(* IEC 61131-3 sources: 2026_Projet_YGO_ExcavatriceDragage/ARCHIVES/Code/SUPERVISION, 3 files *)

(* ---- ST_Safety_Emergency_HmiCmd.st ---- *)
(* ==============================================================
   [IHM] ST_Safety_Emergency_HmiCmd -- Commandes IHM pour la chaine AU
   --------------------------------------------------------------
   Role : structure d'echange pour les commandes operateur
          de la chaine d'arret d'urgence (miroir ST_ModesCmd).
   Pattern : identique a GVL_IHM.Modes.Cmd dans le projet reel.
          L'IHM ecrit ces champs, le programme les consomme.
   ==============================================================
    Docs : DOC/AF/AF_Partie-01_Analyse_Fonctionnelle_v2.0.md
           DOC/AF/AF_Partie-07_Interface_IHM_v2.0.md
*)

TYPE ST_Safety_Emergency_HmiCmd :
STRUCT
    BtnEmergencyArming   : BOOL;   // Front demande rearmement contacteur
    BtnEmergencyCutOff   : BOOL;   // Niveau coupure IHM maintenue
    BtnFaultReset        : BOOL;   // Front acquittement defauts
END_STRUCT
END_TYPE

(* ---- ST_Safety_Emergency_HmiState.st ---- *)
(* ==============================================================
   [IHM] ST_Safety_Emergency_HmiState -- Retours d'etat IHM pour chaine AU
   --------------------------------------------------------------
   Role : structure d'echange pour les retours d'etat de la
          chaine d'arret d'urgence (miroir ST_ModesState).
   Pattern : identique a GVL_IHM.Modes.State dans le projet reel.
          Le programme ecrit ces champs, l'IHM les lit.
   ==============================================================
    Docs : DOC/AF/AF_Partie-01_Analyse_Fonctionnelle_v2.0.md
           DOC/AF/AF_Partie-07_Interface_IHM_v2.0.md
*)

TYPE ST_Safety_Emergency_HmiState :
STRUCT
    // [OK] Etats generaux
    ChainOk              : BOOL;   // Boucle AU fermee (saine)
    ContactorOk          : BOOL;   // Contacteur puissance engage
    PowerCutOffActive    : BOOL;   // Coupure puissance demandee par une safety metier

    // [AU] Sequence de rearmement
    Armable              : BOOL;   // Pret au rearmement (chain OK + pas de lockout + pas de defaut)
    ArmingBusy           : BOOL;   // Sequence armement en cours
    Step                 : INT;    // Etape sequence (0=IDLE, 1=TestA, 2=RestoreA, 3=TestB, 4=RestoreB, 5=Pulse, 6=Confirm)

    // [KO] Diagnostics
    Error                : BOOL;   // Synthese defaut
    ErrorId              : WORD;   // bit0=RedundancyTestFailed, bit1=ArmingFailed
    RedundancyTestFailed : BOOL;   // Auto-test A/B a echoue (canal colle/shunte)
    ArmingFailed         : BOOL;   // Rearmement echoue (timeout confirmation)
    LockoutActive        : BOOL;   // Verrouillage 5s entre tentatives
END_STRUCT
END_TYPE

(* ---- GVL_IHM_AU.st ---- *)
(* ==============================================================
   [IHM] GVL_IHM_AU -- Interface IHM pour le test de la chaine AU
   --------------------------------------------------------------
   Role : point d'echange unique entre l'IHM (Watch/visu) et
          le programme de test de la chaine d'arret d'urgence.
   Pattern : identique a GVL_IHM.Modes (Cmd + State) dans le
          projet reel.
   Usage :
     GVL_IHM_AU.Cmd.BtnEmergencyArming   -> ecrit par l'IHM
     GVL_IHM_AU.State.ContactorOk         -> lu par l'IHM
   ==============================================================
    Docs : DOC/AF/AF_Partie-01_Analyse_Fonctionnelle_v2.0.md
           DOC/AF/AF_Partie-07_Interface_IHM_v2.0.md
*)

{attribute 'qualified_only'}
VAR_GLOBAL
    Cmd   : ST_Safety_Emergency_HmiCmd;    // [IHM] Commandes operateur (Write)
    State : ST_Safety_Emergency_HmiState;  // [IHM] Retours d'etat (Read)
END_VAR
